(* IEC 61131-3 sources: Lasal-MCP/examples/SampleSource/LASALScreenAdvancedSolution/LASALScreenAdvancedSolution/LASALScreenAdvacnedSolution/Stations/Terminal/HMI/Network/MyIONet, 1 file *)

(* ---- ONE_MyIONet_Table.st ---- *)
#define OBJECTS_CONFIG

//Define part of class InputMyIO
#define CROSSHAIR_LENGTH 20
#define CROSSHAIR_WIDTH 1
#define OFFSET_X 10
#define OFFSET_Y 5

FUNCTION GLOBAL TAB ONE_MyIONet
-1$UINT, 0$UINT,
0$UINT, 0$UINT,

6$UDINT,
TO_UDINT(2980745877), "_MyIO", 0$UINT, 3$UINT, 0$UINT,
TO_UDINT(2798398088), "CirleMyIO", 0$UINT, 0$UINT, 1$UINT,
TO_UDINT(3621868871), "InputMyIO", 0$UINT, 0$UINT, 1$UINT,
TO_UDINT(2672428609), "MyColorBar", 0$UINT, 0$UINT, 1$UINT,
TO_UDINT(2517122451), "MyFirstMyIO", 0$UINT, 0$UINT, 1$UINT,
TO_UDINT(2861140242), "UseImageScheme", 0$UINT, 0$UINT, 1$UINT,

_NO_ATTR, TO_UDINT(1612261519), "CIRLEMYIO1",

_NO_ATTR, TO_UDINT(1806949073), "INPUTMYIO1",

_NO_ATTR, TO_UDINT(2191054007), "MYCOLORBAR1",

_NO_ATTR, TO_UDINT(3930858868), "MYFIRSTMYIO1",

_NO_ATTR, TO_UDINT(1892620150), "USEIMAGESCHEME1",

//Internal connections
0$UDINT,
0$UDINT,
0$UDINT,
0$UDINT,

//Initialization values
0$UDINT,
5$UDINT,
TO_UDINT(0), "XPos", TO_UDINT(60),//|MyIONet.CirleMyIO1.XPos;
TO_UDINT(0), "YPos", TO_UDINT(60),//|MyIONet.CirleMyIO1.YPos;
TO_UDINT(0), "CircleRadius", TO_UDINT(80),//|MyIONet.CirleMyIO1.CircleRadius;
TO_UDINT(0), "CircleAngle", TO_UDINT(3600),//|MyIONet.CirleMyIO1.CircleAngle;
TO_UDINT(4), "DelayTime", TO_UDINT(500),//|MyIONet.UseImageScheme1.DelayTime;

//Symbolic initialization values
0$UDINT,
0$UDINT,

//Initialization of string values
0$UDINT,
0$UDINT,

//Configuration of tasks (RealTime, Cyclic, Background)
0$UDINT,
0$UDINT,

0$UDINT,
0$UDINT,

0$UDINT,
0$UDINT,

//External connections
0$UDINT,
5$UDINT,
TO_UDINT(0), "Lse", C_DIR, TO_UDINT(299963966), "Lse","Lse",
TO_UDINT(1), "Lse", C_DIR, TO_UDINT(299963966), "Lse","Lse",
TO_UDINT(2), "Lse", C_DIR, TO_UDINT(299963966), "Lse","Lse",
TO_UDINT(3), "Lse", C_DIR, TO_UDINT(299963966), "Lse","Lse",
TO_UDINT(4), "Lse", C_DIR, TO_UDINT(299963966), "Lse","Lse",

//Magic internal connections
0$UDINT,
0$UDINT,

//Configuration of timeslots of tasks (RealTime, Cyclic)
#ifdef __LSLLDR_TIMESLOTS__
0$UDINT,
0$UDINT,

0$UDINT,
0$UDINT,

#endif //__LSLLDR_TIMESLOTS__

//MultiMaster connections
#ifdef __LSLLDR_MULTIMASTER__
0$UDINT,
0$UDINT,
#endif //__LSLLDR_MULTIMASTER__

//Configuration for task ID (RealTime, CyclicTime)
#ifdef __LSLLDR_TASKID__
"\\\\TASKS2  "
0$UDINT,
0$UDINT,

0$UDINT,
0$UDINT,

0$UDINT,
0$UDINT,

#endif //__LSLLDR_TASKID__

END_FUNCTION
